(* IEC 61131-3 sources: 2026_Projet_YGO_ExcavatriceDragage/CODE_BACKUP/CODE_20260807_v0.5.25/CYCLE, 6 files *)

(* ---- E_CycleStep.st ---- *)
(* ═══════════════════════════════════════════════════════════════
   🔄 E_CycleStep — Étapes de la machine d'état du cycle automatique
   ───────────────────────────────────────────────────────────────
   📄 Doc : DOC/AF_Partie-04_Mode_SemiAuto_Sequenceur_v2.0.md §1
   ═══════════════════════════════════════════════════════════════ *)

TYPE E_CycleStep :
(
  INIT                 := 0,   (* Vérifs cohérence états + sécurités, mise en position init *)
  WORK_POS_SELECT      := 1,   (* Choix opérateur pos travail 1/2 + déplacement validé joystick *)
  DESCENDING_OPEN      := 2,   (* Plongée benne déjà ouvert, M1+M2 synchro *)
  BOTTOM_TOUCH_WAIT    := 3,   (* Attente info BOOL capteur "fond touché" *)
  SYNCHRO_ADJUST       := 4,   (* Désynchro M2 petite vitesse (offset X) → fermeture benne *)
  CTRL_ASCENDING       := 5,   (* Remontée lente de contrôle (vérification fermeture) *)
  ASCENDING_LOADED     := 6,   (* Remontée pleine vitesse charge *)
  DRAINING_PAUSE       := 7,   (* Égouttage temporisé (durée RETAIN) *)
  TRANSLATION_MOVE         := 8,   (* Déplacement translation M3 vers trémie *)
  DESCENDING_OPEN_DUMP := 9,   (* Descente de vidage + ouverture benne *)
  RETURN_WORK_POS      := 10,  (* Retour position travail (remontée synchro) *)
  READY                := 11,  (* Cycle terminé, prêt à reboucler *)
  ERROR_HOLD           := 12   (* Arrêt sûr figé sur défaut (SafeStop) *)
);
END_TYPE

(* ---- E_DiveSearchState.st ---- *)
(* ═══════════════════════════════════════════════════════════════
   🌊 E_DiveSearchState — Phases internes de recherche du fond Kobold
   📄 Doc : DOC/AF_Partie-04_Mode_SemiAuto_Sequenceur_v2.0.md §3ter
   ═══════════════════════════════════════════════════════════════ *)
TYPE E_DiveSearchState :
(
    WAIT_PRECONDITIONS := 0, (* Attente benne ouverte, positions et Kobold au repos *)
    READY_TO_DESCEND   := 1, (* Prêt à assister une demande de descente *)
    SEARCHING_IMMERSION := 2, (* Descente : attente front 0→1 dans fenêtre eau *)
    SEARCHING_BOTTOM    := 3, (* Immersion validée : attente front 1→0 au fond *)
    BOTTOM_CONFIRMED    := 4, (* Fond validé ; extraction peut être demandée *)
    ERROR_HOLD          := 5  (* Séquence invalide, descente assistée interdite *)
);
END_TYPE

(* ---- E_ExtractionSequenceState.st ---- *)
(* ═══════════════════════════════════════════════════════════════
   ⛏️ E_ExtractionSequenceState — Phases extraction assistée
   📄 Doc : DOC/AF_Partie-04_Mode_SemiAuto_Sequenceur_v2.0.md §3ter
   ═══════════════════════════════════════════════════════════════ *)
TYPE E_ExtractionSequenceState :
(
    WAIT_BOTTOM_CONFIRMATION := 0, (* Attente fond Kobold ou attestation opérateur *)
    READY_TO_CLOSE            := 1, (* Prêt à fermer la benne *)
    CLOSING_BUCKET            := 2, (* FB_Bucket ferme M2 seul *)
    CONTROL_ASCENT            := 3, (* M1/M2 synchronisés au palier sans contacteur vitesse *)
    NOMINAL_ASCENT            := 4, (* Montée couplée avec vitesse demandée opérateur *)
    ERROR_HOLD                := 5  (* Défaut extraction, reprise interdite avant reset *)
);
END_TYPE

(* ---- FB_Cycle.st ---- *)
(* ═══════════════════════════════════════════════════════════════
   🔄 FB_Cycle — Séquenceur du Cycle Automatique (Grafcet de dragage)
   ───────────────────────────────────────────────────────────────
   📄 Doc : DOC/AF_Partie-04_Mode_SemiAuto_Sequenceur_v2.0.md
   🔌 Conforme au contrat FB standard (Partie3 §1bis).
   ═══════════════════════════════════════════════════════════════ *)

FUNCTION_BLOCK FB_Cycle
VAR_INPUT
    Enable                  : BOOL;         // Activation générale du séquenceur
    Reset                   : BOOL;         // Acquittement défaut (front)
    PowerContactorEngaged   : BOOL;         // Chaîne de sécurité OK
    CycleMotionPermit       : BOOL;         // Homme-mort + joystick actif
    HeartbeatIhmOk          : BOOL;         // 💓 IHM↔PLC valide ; FALSE = repli cycle obligatoire

    // Commandes opérateur
    StartCycle              : BOOL;         // Demande lancement / reprise cycle (IHM)
    PauseCycle              : BOOL;         // Demande pause temporaire (IHM)
    AbortCycle              : BOOL;         // Demande abandon cycle (IHM)

    // Cibles et paramètres
    SetDepthM               : REAL;         // Profondeur de consigne (négative)
    SetOffsetM              : REAL;         // Écart de fermeture benne cible
    SelectedTargetNum_IHM   : INT;          // Cible sélectionnée (2=P2, 3=P1)

    // Feedbacks physique & matériel
    KoboldContactFond       : BOOL;         // Retour dédié Kobold : TRUE = contact fond détecté
    LimitLegalReached       : BOOL;         // Limite légale atteinte (descente interdite)
    LimitLegalDepthM        : REAL;         // Profondeur légale minimale autorisée
    WinchSyncError          : BOOL;         // Désynchronisme bloquant M1/M2
    WinchSyncDeltaM         : REAL;         // Écart codeurs M1/M2 pour diagnostic
    M1_CablePosM            : REAL;         // Position câble treuil M1 (recalée)
    M2_CablePosM            : REAL;         // Position câble treuil M2 (recalée)
    M1_MeasuredSpeedMps     : REAL;         // Vitesse linéaire mesurée M1 (m/s)
    M2_MeasuredSpeedMps     : REAL;         // Vitesse linéaire mesurée M2 (m/s)
    SpeedMismatchThresholdMps : REAL;       // Seuil écart vitesse ; 0 = contrôle désactivé
    SpeedMismatchTimeout    : TIME;         // Durée de confirmation ; 0 = contrôle désactivé
    CableLimitM1AscentM     : REAL;         // Limite haute d'exploitation M1 ; seuil de fin ASCENDING_LOADED

    // Feedbacks Translation M3
    Translation_At_P1           : BOOL;     // Capteur position P1 (ex-Fosse1)
    Translation_At_P2           : BOOL;     // Capteur position P2 (ex-Fosse2)
    Translation_At_Maintenance  : BOOL;     // Capteur fin de course maintenance
    Translation_At_Tremie       : BOOL;     // Capteur fin de course trémie
    Translation_Busy            : BOOL;     // Mouvement translation en cours
    Translation_Done            : BOOL;     // Cible translation atteinte

    // Feedbacks Benne
    Benne_Busy              : BOOL;         // Mouvement mâchoires benne en cours
    Benne_Done              : BOOL;         // Mouvement ouverture/fermeture terminé
    Benne_IsOpen            : BOOL;         // Benne mécaniquement ouvert mémorisé
    Benne_IsClosed          : BOOL;         // Benne mécaniquement fermé mémorisé
END_VAR
VAR_OUTPUT
    Ready                   : BOOL;         // Séquenceur disponible
    Busy                    : BOOL;         // Cycle automatique actif
    Done                    : BOOL;         // Cycle automatique complété
    Error                   : BOOL;         // Défaut cycle
    ErrorId                 : WORD;         // bit0: Timeout/limite, bit1: désynchronisme, bit2: cible invalide, bit3: stabilisation impossible, bit4: écart vitesse, bit5: perte heartbeat
    SpeedMismatchMps        : REAL;         // Écart absolu vitesse M1/M2 (m/s)
    SpeedMismatchActive     : BOOL;         // Seuil vitesse dépassé sur le cycle courant
    SpeedMismatchConfirmed  : BOOL;         // Écart vitesse confirmé pendant SpeedMismatchTimeout

    // Commandes structurées (demandes de mouvement)
    WinchM1Cmd              : ST_WinchCmdDemand;        // Demande treuil M1
    WinchM2Cmd              : ST_WinchCmdDemand;        // Demande treuil M2
    TranslationCmd          : ST_TranslationCmdDemand;  // Demande translation M3
    BucketCmd               : ST_BucketCmdDemand;       // Demande benne

    // Métadonnées d'affichage IHM
    CycleStep               : E_CycleStep;  // Étape active du Grafcet
    CycleStateStr           : STRING(80);   // Libellé en clair de l'étape
END_VAR
VAR
    ResetEdge               : R_TRIG;
    StartEdge               : R_TRIG;
    PauseEdge               : R_TRIG;
    AbortEdge               : R_TRIG;

    // Séquencement
    State                   : E_CycleStep := E_CycleStep.INIT;
    SavedState              : E_CycleStep := E_CycleStep.INIT;
    IsPaused                : BOOL := FALSE;

    // Mémorisations et Timers
    TouchPositionM          : REAL;         // Position M1 mémorisée lors du contact fond
    RaiseTargetM            : REAL;         // Profondeur de remontée mémorisée
    DrainingTimer           : TON;          // Temporisateur de vidage (égouttage)
    StabilizationTimer      : TON;          // Temporisation maximale de remontée lente après fermeture
    SpeedMismatchTimer      : TON;          // Confirmation temporelle écart de vitesse M1/M2
    SelectedWorkTarget      : INT;          // Cible de travail mémorisée (2=P2 ou 3=P1)

    // Paramètres internes
    CtrlAscentDistM         : REAL := 2.0;      // Distance de remontée lente de contrôle
    CtrlAscentToleranceM    : REAL := 0.25;     // Écart maximal admis entre les deux codeurs
    CtrlAscentTimeout       : TIME := T#30s;    // Temps maximal pour atteindre la zone de stabilisation
    DrainingTime            : TIME := T#5s;     // Temps d'égouttage par défaut
END_VAR

// === IMPLEMENTATION ===

// 🛑 1. GATES DE SÉCURITÉ ET BLOCAGE
IF NOT Enable OR NOT PowerContactorEngaged THEN
    WinchM1Cmd.StartStop   := FALSE;
    WinchM1Cmd.Direction   := 0;
    WinchM1Cmd.SpeedPct    := 0.0;

    WinchM2Cmd.StartStop   := FALSE;
    WinchM2Cmd.Direction   := 0;
    WinchM2Cmd.SpeedPct    := 0.0;

    TranslationCmd.Start   := FALSE;
    TranslationCmd.Target  := 0;

    BucketCmd.Open         := FALSE;
    BucketCmd.Close        := FALSE;
    BucketCmd.KoboldContactorCmd := FALSE;

    State                := E_CycleStep.INIT;
    CycleStep            := E_CycleStep.INIT;
    CycleStateStr        := 'ARRÊT : SÉCURITÉ ABSENTE OU AUTO DÉSACTIVÉ';
    Ready                := FALSE;
    Busy                 := FALSE;
    Done                 := FALSE;
    RETURN;
END_IF;

Ready := TRUE;
ResetEdge(CLK := Reset);
StartEdge(CLK := StartCycle);
PauseEdge(CLK := PauseCycle);
AbortEdge(CLK := AbortCycle);

// ⏱️ T36 — surveillance indépendante de la remontée lente : un codeur bloqué
// ne doit jamais laisser le cycle attendre indéfiniment.
StabilizationTimer(IN := (State = E_CycleStep.CTRL_ASCENDING), PT := CtrlAscentTimeout);

// 📏 T43 — comparaison vitesse réelle M1/M2.
SpeedMismatchMps := ABS(M1_MeasuredSpeedMps - M2_MeasuredSpeedMps);
SpeedMismatchActive := (State = E_CycleStep.CTRL_ASCENDING)
                       AND CycleMotionPermit
                       AND (SpeedMismatchThresholdMps > 0.0)
                       AND (SpeedMismatchTimeout > T#0ms)
                       AND (SpeedMismatchMps > SpeedMismatchThresholdMps);
SpeedMismatchTimer(IN := SpeedMismatchActive, PT := SpeedMismatchTimeout);
SpeedMismatchConfirmed := SpeedMismatchTimer.Q;

IF ResetEdge.Q THEN
    Error := FALSE;
    ErrorId := 16#0000;
    IsPaused := FALSE;
    SavedState := E_CycleStep.INIT;
    IF State = E_CycleStep.ERROR_HOLD THEN
        State := E_CycleStep.INIT;
    END_IF;
END_IF;

// 💓 Perte IHM : repli mémorisé. La reconnexion seule ne relance jamais le cycle.
IF NOT HeartbeatIhmOk AND State <> E_CycleStep.ERROR_HOLD THEN
    Error := TRUE;
    ErrorId := ErrorId OR 16#0020;
    State := E_CycleStep.ERROR_HOLD;
END_IF;

// Défaut de synchronisme : arrêt sûr et acquittement obligatoire.
IF WinchSyncError AND State <> E_CycleStep.ERROR_HOLD THEN
    Error := TRUE;
    ErrorId := ErrorId OR 16#0002;
    State := E_CycleStep.ERROR_HOLD;
END_IF;

// 🛡️ T43 — écart de vitesse confirmé : arrêt du cycle et ERROR_HOLD.
IF SpeedMismatchConfirmed AND State <> E_CycleStep.ERROR_HOLD THEN
    Error := TRUE;
    ErrorId := ErrorId OR 16#0010;
    State := E_CycleStep.ERROR_HOLD;
END_IF;

// Gestion de la Pause
IF PauseEdge.Q AND Busy AND NOT IsPaused THEN
    IsPaused := TRUE;
    SavedState := State;
    State := E_CycleStep.ERROR_HOLD; // Fige les mouvements
ELSIF StartEdge.Q AND IsPaused THEN
    IsPaused := FALSE;
    State := SavedState; // Reprise à l'étape sauvegardée
END_IF;

// Gestion de l'Abandon
IF AbortEdge.Q THEN
    IsPaused := FALSE;
    State := E_CycleStep.INIT;
END_IF;

// 🔁 2. LOGIQUE DU SÉQUENCEUR (Machine d'état)
CASE State OF

    E_CycleStep.INIT:
        CycleStep := E_CycleStep.INIT;
        CycleStateStr := 'VÉRIFICATION COHÉRENCE SYSTÈME';

        WinchM1Cmd.StartStop := FALSE;
        WinchM1Cmd.Direction := 0;
        WinchM1Cmd.SpeedPct  := 0.0;

        WinchM2Cmd.StartStop := FALSE;
        WinchM2Cmd.Direction := 0;
        WinchM2Cmd.SpeedPct  := 0.0;

        TranslationCmd.Start := FALSE;
        TranslationCmd.Target := 0;

        BucketCmd.Open  := FALSE;
        BucketCmd.Close := FALSE;
        BucketCmd.KoboldContactorCmd := FALSE;

        Busy  := FALSE;
        Done  := FALSE;

        // Transition si système sain et réarmé (front reset ou démarrage)
        IF StartEdge.Q THEN
            State := E_CycleStep.WORK_POS_SELECT;
        END_IF;

    E_CycleStep.WORK_POS_SELECT:
        CycleStep := E_CycleStep.WORK_POS_SELECT;
        CycleStateStr := 'SÉLECTION POSITION TRAVAIL (FOSSE 1 / 2)';
        Busy := TRUE;

        // Choix cible — P2/P1 (cibles 2/3)
        IF (SelectedTargetNum_IHM <> 2) AND (SelectedTargetNum_IHM <> 3) THEN
            Error := TRUE;
            ErrorId := ErrorId OR 16#0004;
            State := E_CycleStep.ERROR_HOLD;
        ELSIF SelectedTargetNum_IHM = 2 OR SelectedTargetNum_IHM = 3 THEN
            SelectedWorkTarget := SelectedTargetNum_IHM;
            TranslationCmd.Target := SelectedWorkTarget;
            TranslationCmd.Start := CycleMotionPermit;

            // Attente positionnement translation
            IF CycleMotionPermit AND ((SelectedWorkTarget = 2 AND Translation_At_P2)
               OR (SelectedWorkTarget = 3 AND Translation_At_P1)) THEN
                TranslationCmd.Start := FALSE;
                State := E_CycleStep.DESCENDING_OPEN;
            END_IF;
        END_IF;

    E_CycleStep.DESCENDING_OPEN:
        CycleStep := E_CycleStep.DESCENDING_OPEN;
        CycleStateStr := 'PLONGÉE BENNE OUVERT';

        // M1 et M2 descendent ensemble (synchro gérée en aval)
        WinchM1Cmd.StartStop := TRUE;
        WinchM1Cmd.Direction := -1;
        WinchM1Cmd.SpeedPct  := 50.0;

        WinchM2Cmd.StartStop := TRUE;
        WinchM2Cmd.Direction := -1;
        WinchM2Cmd.SpeedPct  := 50.0;

        BucketCmd.KoboldContactorCmd := TRUE;

        // Transition uniquement sur le retour dédié Kobold.
        IF CycleMotionPermit AND KoboldContactFond THEN
            WinchM1Cmd.StartStop := FALSE;
            WinchM2Cmd.StartStop := FALSE;
            BucketCmd.KoboldContactorCmd := FALSE;
            TouchPositionM := M1_CablePosM;
            IF LimitLegalDepthM < -0.01 THEN
                RaiseTargetM := MAX(TouchPositionM + 0.5, LimitLegalDepthM + 0.5);
            ELSE
                RaiseTargetM := TouchPositionM + 0.5;
            END_IF;
            State := E_CycleStep.BOTTOM_TOUCH_WAIT;
        ELSIF LimitLegalReached THEN
            Error := TRUE;
            ErrorId := ErrorId OR 16#0001;
            WinchM1Cmd.StartStop := FALSE;
            WinchM2Cmd.StartStop := FALSE;
            BucketCmd.KoboldContactorCmd := FALSE;
            State := E_CycleStep.ERROR_HOLD;
        END_IF;

    E_CycleStep.BOTTOM_TOUCH_WAIT:
        CycleStep := E_CycleStep.BOTTOM_TOUCH_WAIT;
        CycleStateStr := 'REMONTÉE SÉCURISÉE APRÈS CONTACT FOND';

        WinchM1Cmd.StartStop := TRUE;
        WinchM1Cmd.Direction := 1;
        WinchM1Cmd.SpeedPct := 20.0;

        WinchM2Cmd.StartStop := TRUE;
        WinchM2Cmd.Direction := 1;
        WinchM2Cmd.SpeedPct := 20.0;

        // Les deux treuils restent synchronisés jusqu'au-dessus de la limite légale.
        IF CycleMotionPermit AND (M1_CablePosM >= RaiseTargetM) AND (M2_CablePosM >= RaiseTargetM) THEN
            WinchM1Cmd.StartStop := FALSE;
            WinchM2Cmd.StartStop := FALSE;
            State := E_CycleStep.SYNCHRO_ADJUST;
        END_IF;

    E_CycleStep.SYNCHRO_ADJUST:
        CycleStep := E_CycleStep.SYNCHRO_ADJUST;
        CycleStateStr := 'FERMETURE DU GODET / EXCAVATION';

        WinchM1Cmd.StartStop := FALSE;

        // Déclenchement fermeture benne
        BucketCmd.Close := TRUE;

        // Transition si benne fermé avec succès
        IF CycleMotionPermit AND Benne_Done AND Benne_IsClosed THEN
            BucketCmd.Close := FALSE;
            State := E_CycleStep.CTRL_ASCENDING;
        END_IF;

    E_CycleStep.CTRL_ASCENDING:
        CycleStep := E_CycleStep.CTRL_ASCENDING;
        CycleStateStr := 'REMONTÉE LENTE DE CONTRÔLE';

        // M1 et M2 montent lentement en synchro
        WinchM1Cmd.StartStop := TRUE;
        WinchM1Cmd.Direction := 1;
        WinchM1Cmd.SpeedPct  := 20.0;

        WinchM2Cmd.StartStop := TRUE;
        WinchM2Cmd.Direction := 1;
        WinchM2Cmd.SpeedPct  := 20.0;

        // Contrôle des deux codeurs
        IF WinchSyncError OR (ABS(M1_CablePosM - M2_CablePosM) > CtrlAscentToleranceM) THEN
            Error := TRUE;
            ErrorId := ErrorId OR 16#0008;
            State := E_CycleStep.ERROR_HOLD;
        ELSIF CycleMotionPermit
           AND (M1_CablePosM >= (TouchPositionM + CtrlAscentDistM))
           AND (M2_CablePosM >= (TouchPositionM + CtrlAscentDistM))
           AND (ABS(M1_CablePosM - M2_CablePosM) <= CtrlAscentToleranceM) THEN
            State := E_CycleStep.ASCENDING_LOADED;
        ELSIF StabilizationTimer.Q THEN
            Error := TRUE;
            ErrorId := ErrorId OR 16#0008;
            State := E_CycleStep.ERROR_HOLD;
        END_IF;

    E_CycleStep.ASCENDING_LOADED:
        CycleStep := E_CycleStep.ASCENDING_LOADED;
        CycleStateStr := 'REMONTÉE EN CHARGE';

        WinchM1Cmd.StartStop := TRUE;
        WinchM1Cmd.Direction := 1;
        WinchM1Cmd.SpeedPct  := 70.0;

        WinchM2Cmd.StartStop := TRUE;
        WinchM2Cmd.Direction := 1;
        WinchM2Cmd.SpeedPct  := 70.0;

        // Transition alignée sur la limite haute d'exploitation
        IF CycleMotionPermit AND M1_CablePosM >= CableLimitM1AscentM THEN
            WinchM1Cmd.StartStop := FALSE;
            WinchM2Cmd.StartStop := FALSE;
            State := E_CycleStep.DRAINING_PAUSE;
        END_IF;

    E_CycleStep.DRAINING_PAUSE:
        CycleStep := E_CycleStep.DRAINING_PAUSE;
        CycleStateStr := 'ÉGOUTTAGE DU GODET EN COURS';

        WinchM1Cmd.StartStop := FALSE;
        WinchM2Cmd.StartStop := FALSE;

        DrainingTimer(IN := TRUE, PT := DrainingTime);
        IF CycleMotionPermit AND DrainingTimer.Q THEN
            DrainingTimer(IN := FALSE);
            State := E_CycleStep.TRANSLATION_MOVE;
        END_IF;

    E_CycleStep.TRANSLATION_MOVE:
        CycleStep := E_CycleStep.TRANSLATION_MOVE;
        CycleStateStr := 'DÉPLACEMENT VERS TRÉMIE DE VIDANGE';

        TranslationCmd.Target := 1; // Trémie
        TranslationCmd.Start := TRUE;

        // Transition si translation arrivé à la trémie
        IF CycleMotionPermit AND Translation_At_Tremie THEN
            TranslationCmd.Start := FALSE;
            State := E_CycleStep.DESCENDING_OPEN_DUMP;
        END_IF;

    E_CycleStep.DESCENDING_OPEN_DUMP:
        CycleStep := E_CycleStep.DESCENDING_OPEN_DUMP;
        CycleStateStr := 'VIDANGE / OUVERTURE DU GODET';

        BucketCmd.Open := TRUE;

        // Transition si benne ouvert avec succès
        IF CycleMotionPermit AND Benne_Done AND Benne_IsOpen THEN
            BucketCmd.Open := FALSE;
            State := E_CycleStep.RETURN_WORK_POS;
        END_IF;

    E_CycleStep.RETURN_WORK_POS:
        CycleStep := E_CycleStep.RETURN_WORK_POS;
        CycleStateStr := 'RETOUR VERS FOSSE DE TRAVAIL';

        TranslationCmd.Target := SelectedWorkTarget;
        TranslationCmd.Start := TRUE;

        // Transition si translation de retour sur sa position de travail
        IF CycleMotionPermit AND ((SelectedWorkTarget = 2 AND Translation_At_P2)
           OR (SelectedWorkTarget = 3 AND Translation_At_P1)) THEN
            TranslationCmd.Start := FALSE;
            State := E_CycleStep.READY;
        END_IF;

    E_CycleStep.READY:
        CycleStep := E_CycleStep.READY;
        CycleStateStr := 'CYCLE AUTOMATIQUE COMPLÉTÉ - PRÊT';

        WinchM1Cmd.StartStop := FALSE;
        WinchM2Cmd.StartStop := FALSE;
        TranslationCmd.Start := FALSE;
        Done  := TRUE;
        Busy  := FALSE;

        // Rebouclage manuel ou auto sur Start
        IF StartEdge.Q THEN
            Done := FALSE;
            State := E_CycleStep.DESCENDING_OPEN;
        END_IF;

    E_CycleStep.ERROR_HOLD:
        CycleStep := E_CycleStep.ERROR_HOLD;
        CycleStateStr := 'CYCLE SUSPENDU (PAUSE OU ARRÊT DE SÉCURITÉ)';

        WinchM1Cmd.StartStop := FALSE;
        WinchM2Cmd.StartStop := FALSE;
        TranslationCmd.Start := FALSE;

        BucketCmd.Open  := FALSE;
        BucketCmd.Close := FALSE;

END_CASE;

// 🛑 Relâchement homme-mort : aucune demande d'actionneur ne reste active.
// L'étape est mémorisée et reprend au prochain appui valide.
IF Busy AND NOT CycleMotionPermit THEN
    WinchM1Cmd.StartStop := FALSE;
    WinchM2Cmd.StartStop := FALSE;
    TranslationCmd.Start := FALSE;
    BucketCmd.Open := FALSE;
    BucketCmd.Close := FALSE;
    BucketCmd.KoboldContactorCmd := FALSE;
END_IF;

END_FUNCTION_BLOCK

(* ---- FB_DiveSearch.st ---- *)
(* ═══════════════════════════════════════════════════════════════
   🌊 FB_DiveSearch — Assistance plongée et recherche du fond Kobold
   ───────────────────────────────────────────────────────────────
   📄 Doc : DOC/AF_Partie-04_Mode_SemiAuto_Sequenceur_v2.0.md §3ter
   🛡️ Sécurité : T81/T82. Jamais de descente assistée sans séquence 0→1→0 valide.
   🧩 Responsabilité : qualifie le Kobold et autorise uniquement la descente cohérente.
   🔌 Interface : intention de descente + mesures → autorisation + fond validé.
   ═══════════════════════════════════════════════════════════════ *)
FUNCTION_BLOCK FB_DiveSearch
VAR_INPUT
    Enable                 : BOOL;
    Reset                  : BOOL;
    PowerContactorEngaged        : BOOL;
    Mode                   : E_Mode;
    MotionRequestActive    : BOOL; (* Intention déjà arbitrée en amont *)
    MotionDirection        : INT;  (* -1 = descente *)
    BucketIsOpen           : BOOL;
    KoboldImmersed         : BOOL; (* FALSE hors eau/fond ; TRUE immergé *)
    M1Position_M           : REAL;
    M2Position_M           : REAL;
    PositionsValid         : BOOL;
    DiveStartMin_M         : REAL;
    ImmersionUpper_M       : REAL;
    ImmersionLower_M       : REAL;
    // 🆕 2026-08-07 (14) — retour terrain, demande explicite : réglages DiveStartMin_M/
    // ImmersionUpper_M/ImmersionLower_M pas encore calibrés sur site, bloquaient WAIT_PRECONDITIONS
    // (bit2 config) sans aucun moyen de progresser dans la séquence pendant les essais. Si TRUE,
    // saute entièrement ErrorCausePresent (bit2) ET le test WAIT_PRECONDITIONS -- transition directe
    // vers READY_TO_DESCEND. Défaut FALSE : comportement standard inchangé.
    BypassPreconditions    : BOOL := FALSE;
END_VAR
VAR_OUTPUT
    Ready                  : BOOL;
    Busy                   : BOOL;
    Done                   : BOOL;
    Error                  : BOOL;
    ErrorId                : WORD; (* bit0: préconditions, bit1: séquence Kobold invalide, bit2: configuration seuils invalide *)
    State                  : E_State;
    StateAtError           : E_State;
    DiveState              : E_DiveSearchState;
    DescendPermit          : BOOL; (* Autorise uniquement la demande de descente active *)
    KoboldMeasureEnable    : BOOL;
    BottomTouchConfirmed   : BOOL;
    OperatorActionId       : WORD;
    OperatorAction         : STRING(120);
END_VAR
VAR
    ResetEdge              : R_TRIG;
    KoboldRiseEdge         : R_TRIG;
    KoboldFallEdge         : F_TRIG;
    ImmersionConfirmed     : BOOL;
    ErrorCausePresent      : BOOL;
END_VAR

IF NOT Enable OR NOT PowerContactorEngaged THEN
    Ready := FALSE; Busy := FALSE; Done := FALSE;
    DescendPermit := FALSE; KoboldMeasureEnable := FALSE;
    BottomTouchConfirmed := FALSE;
    State := E_State.DISABLED;
    StateAtError := E_State.DISABLED;
    DiveState := E_DiveSearchState.WAIT_PRECONDITIONS;
    OperatorActionId := 0; OperatorAction := '';
    ImmersionConfirmed := FALSE;
    RETURN;
END_IF;

ResetEdge(CLK := Reset);
KoboldRiseEdge(CLK := KoboldImmersed);
KoboldFallEdge(CLK := KoboldImmersed);

ErrorCausePresent := NOT BypassPreconditions AND ((DiveStartMin_M < ImmersionUpper_M)
                  OR (ImmersionUpper_M <= ImmersionLower_M));
IF ErrorCausePresent THEN
    ErrorId := ErrorId OR 16#0004;
END_IF;

(* Reset = front + causes disparues ; aucun redémarrage automatique. *)
IF ResetEdge.Q AND NOT ErrorCausePresent AND NOT KoboldImmersed AND NOT MotionRequestActive THEN
    ErrorId := 16#0000;
    ImmersionConfirmed := FALSE;
    BottomTouchConfirmed := FALSE;
    StateAtError := E_State.DISABLED;
    DiveState := E_DiveSearchState.WAIT_PRECONDITIONS;
END_IF;

DescendPermit := FALSE; KoboldMeasureEnable := FALSE;
Ready := FALSE; Busy := FALSE; Done := FALSE;
OperatorActionId := 0; OperatorAction := '';

IF ErrorId <> 16#0000 THEN
    State := E_State.READY;
    DiveState := E_DiveSearchState.ERROR_HOLD;
    OperatorActionId := 16#0180;
    OperatorAction := 'Vérifier les conditions puis réarmer avant une nouvelle plongée.';
ELSE
    CASE DiveState OF
        E_DiveSearchState.WAIT_PRECONDITIONS:
            State := E_State.INIT;
            IF NOT BypassPreconditions
               AND (NOT BucketIsOpen OR NOT PositionsValid OR KoboldImmersed
                    OR (M1Position_M < DiveStartMin_M) OR (M2Position_M < DiveStartMin_M)) THEN
                OperatorActionId := 16#0100;
                OperatorAction := 'Vérifier les conditions initiales de plongée.';
            ELSE
                DiveState := E_DiveSearchState.READY_TO_DESCEND;
            END_IF;

        E_DiveSearchState.READY_TO_DESCEND:
            State := E_State.READY;
            Ready := TRUE;
            OperatorActionId := 16#0101;
            OperatorAction := 'Demander une descente pour rechercher le fond.';
            IF MotionRequestActive AND (MotionDirection = -1) THEN
                DiveState := E_DiveSearchState.SEARCHING_IMMERSION;
            END_IF;

        E_DiveSearchState.SEARCHING_IMMERSION:
            State := E_State.BUSY;
            Busy := TRUE;
            DescendPermit := MotionRequestActive AND (MotionDirection = -1);
            KoboldMeasureEnable := TRUE;
            OperatorActionId := 16#0102;
            OperatorAction := 'Maintenir la descente : recherche immersion Kobold.';
            IF KoboldRiseEdge.Q THEN
                IF (M1Position_M <= ImmersionUpper_M) AND (M1Position_M >= ImmersionLower_M)
                   AND (M2Position_M <= ImmersionUpper_M) AND (M2Position_M >= ImmersionLower_M) THEN
                    ImmersionConfirmed := TRUE;
                    DiveState := E_DiveSearchState.SEARCHING_BOTTOM;
                ELSE
                    ErrorId := ErrorId OR 16#0002;
                    StateAtError := State;
                END_IF;
            ELSIF (M1Position_M < ImmersionLower_M) OR (M2Position_M < ImmersionLower_M) THEN
                ErrorId := ErrorId OR 16#0002;
                StateAtError := State;
            END_IF;

        E_DiveSearchState.SEARCHING_BOTTOM:
            State := E_State.BUSY;
            Busy := TRUE;
            DescendPermit := MotionRequestActive AND (MotionDirection = -1);
            KoboldMeasureEnable := TRUE;
            OperatorActionId := 16#0103;
            OperatorAction := 'Maintenir la descente : immersion validée, recherche du fond.';
            IF KoboldFallEdge.Q AND ImmersionConfirmed THEN
                BottomTouchConfirmed := TRUE;
                ImmersionConfirmed := FALSE;
                DiveState := E_DiveSearchState.BOTTOM_CONFIRMED;
            END_IF;

        E_DiveSearchState.BOTTOM_CONFIRMED:
            State := E_State.DONE;
            Done := TRUE;
            OperatorActionId := 16#0104;
            OperatorAction := 'Fond détecté : demander la fermeture ou l extraction.';

        E_DiveSearchState.ERROR_HOLD:
            State := E_State.READY;
    END_CASE;
END_IF;

Error := (ErrorId <> 16#0000);

(* ---- FB_ExtractionSequence.st ---- *)
(* ═══════════════════════════════════════════════════════════════
   ⛏️ FB_ExtractionSequence — Fermeture benne et remontée assistée
   ───────────────────────────────────────────────────────────────
   📄 Doc : DOC/AF_Partie-04_Mode_SemiAuto_Sequenceur_v2.0.md §3ter
   🛡️ Sécurité : aucune remontée assistée sans fond confirmé ; palier 1 au contrôle.
   🧩 Responsabilité : séquence métier, jamais commande directe de contacteur.
   ═══════════════════════════════════════════════════════════════ *)
FUNCTION_BLOCK FB_ExtractionSequence
VAR_INPUT
    Enable                     : BOOL;
    Reset                      : BOOL;
    PowerContactorEngaged            : BOOL;
    Mode                       : E_Mode;
    MotionRequestActive        : BOOL;
    MotionDirection            : INT; (* +1 = montée *)
    BottomPositionConfirmed    : BOOL;
    BucketIsClosed             : BOOL;
    BucketBusy                 : BOOL;
    BucketError                : BOOL;
    WinchSyncError             : BOOL;
    M1Position_M               : REAL;
    M2Position_M               : REAL;
    M1MeasuredSpeedValid       : BOOL;
    M2MeasuredSpeedValid       : BOOL;
    PositionsValid             : BOOL;
    ControlAscentDistance_M    : REAL;
END_VAR
VAR_OUTPUT
    Ready                      : BOOL;
    Busy                       : BOOL;
    Done                       : BOOL;
    Error                      : BOOL;
    ErrorId                    : WORD; (* bit0: fond absent, bit1: fermeture, bit2: contrôle remontée, bit3: configuration *)
    State                      : E_State;
    StateAtError               : E_State;
    ExtractionState            : E_ExtractionSequenceState;
    BucketCloseRequest         : BOOL;
    AscentPermit               : BOOL;
    ForceMinSpeedStep          : BOOL;
    BottomConfirmationConsumed : BOOL;
    OperatorActionId           : WORD;
    OperatorAction             : STRING(120);
END_VAR
VAR
    ResetEdge                  : R_TRIG;
    ControlStartM1Position_M   : REAL;
    ControlStartM2Position_M   : REAL;
    ErrorCausePresent          : BOOL;
END_VAR

IF NOT Enable OR NOT PowerContactorEngaged THEN
    Ready := FALSE; Busy := FALSE; Done := FALSE;
    BucketCloseRequest := FALSE; AscentPermit := FALSE; ForceMinSpeedStep := FALSE;
    BottomConfirmationConsumed := FALSE;
    State := E_State.DISABLED;
    StateAtError := E_State.DISABLED;
    ExtractionState := E_ExtractionSequenceState.WAIT_BOTTOM_CONFIRMATION;
    OperatorActionId := 0; OperatorAction := '';
    RETURN;
END_IF;

ResetEdge(CLK := Reset);
ErrorCausePresent := (ControlAscentDistance_M <= 0.0);
IF ErrorCausePresent THEN
    ErrorId := ErrorId OR 16#0008;
END_IF;
IF ResetEdge.Q AND NOT ErrorCausePresent AND NOT MotionRequestActive THEN
    ErrorId := 16#0000;
    StateAtError := E_State.DISABLED;
    ExtractionState := E_ExtractionSequenceState.WAIT_BOTTOM_CONFIRMATION;
END_IF;

Ready := FALSE; Busy := FALSE; Done := FALSE;
BucketCloseRequest := FALSE; AscentPermit := FALSE; ForceMinSpeedStep := FALSE;
BottomConfirmationConsumed := FALSE;
OperatorActionId := 0; OperatorAction := '';

IF ErrorId <> 16#0000 THEN
    State := E_State.READY;
    ExtractionState := E_ExtractionSequenceState.ERROR_HOLD;
    OperatorActionId := 16#0280;
    OperatorAction := 'Vérifier la benne et les treuils puis réarmer avant de reprendre.';
ELSE
    CASE ExtractionState OF
        E_ExtractionSequenceState.WAIT_BOTTOM_CONFIRMATION:
            State := E_State.INIT;
            IF BottomPositionConfirmed THEN
                ExtractionState := E_ExtractionSequenceState.READY_TO_CLOSE;
            ELSE
                OperatorActionId := 16#0200;
                OperatorAction := 'Confirmer que la benne est posée au fond avant extraction.';
            END_IF;

        E_ExtractionSequenceState.READY_TO_CLOSE:
            State := E_State.READY;
            Ready := TRUE;
            OperatorActionId := 16#0201;
            OperatorAction := 'Demander la montée pour fermer la benne.';
            IF MotionRequestActive AND (MotionDirection = 1) THEN
                BottomConfirmationConsumed := TRUE;
                ExtractionState := E_ExtractionSequenceState.CLOSING_BUCKET;
            END_IF;

        E_ExtractionSequenceState.CLOSING_BUCKET:
            State := E_State.BUSY;
            Busy := TRUE;
            BucketCloseRequest := MotionRequestActive AND (MotionDirection = 1);
            OperatorActionId := 16#0202;
            OperatorAction := 'Maintenir la montée : fermeture de la benne en cours.';
            IF BucketError THEN
                ErrorId := ErrorId OR 16#0002;
                StateAtError := State;
            ELSIF BucketIsClosed AND NOT BucketBusy THEN
                ControlStartM1Position_M := M1Position_M;
                ControlStartM2Position_M := M2Position_M;
                ExtractionState := E_ExtractionSequenceState.CONTROL_ASCENT;
            END_IF;

        E_ExtractionSequenceState.CONTROL_ASCENT:
            State := E_State.BUSY;
            Busy := TRUE;
            AscentPermit := MotionRequestActive AND (MotionDirection = 1);
            ForceMinSpeedStep := TRUE;
            OperatorActionId := 16#0203;
            OperatorAction := 'Maintenir la montée : contrôle charge au palier minimal.';
            IF WinchSyncError OR NOT PositionsValid OR NOT M1MeasuredSpeedValid OR NOT M2MeasuredSpeedValid THEN
                ErrorId := ErrorId OR 16#0004;
                StateAtError := State;
            ELSIF (M1Position_M >= (ControlStartM1Position_M + ControlAscentDistance_M))
               AND (M2Position_M >= (ControlStartM2Position_M + ControlAscentDistance_M)) THEN
                ExtractionState := E_ExtractionSequenceState.NOMINAL_ASCENT;
            END_IF;

        E_ExtractionSequenceState.NOMINAL_ASCENT:
            State := E_State.BUSY;
            Busy := TRUE;
            AscentPermit := MotionRequestActive AND (MotionDirection = 1);
            OperatorActionId := 16#0204;
            OperatorAction := 'Maintenir la montée : extraction en cours.';
            IF WinchSyncError OR NOT PositionsValid THEN
                ErrorId := ErrorId OR 16#0004;
                StateAtError := State;
            END_IF;

        E_ExtractionSequenceState.ERROR_HOLD:
            State := E_State.READY;
    END_CASE;
END_IF;

Error := (ErrorId <> 16#0000);
